// TIA Portal V17 export
FUNCTION "FC_T02_Bobines" : Void   // FC102, LAD
{ S7_Optimized_Access := 'TRUE' }
// stored: SetENOAutomatically false
   VAR_INPUT
      Entree_1 : Bool;
      Bp_Set : Bool;
      Bp_Reset : Bool;
      Entree_2 : Bool;
   END_VAR
   VAR_OUTPUT
      Sortie_1 : Bool;
      Sortie_2 : Bool;
      Sortie_3 : Bool;
   END_VAR
   VAR_IN_OUT
      Memoire : Bool;
   END_VAR
BEGIN

REGION Network 1: Bobine simple
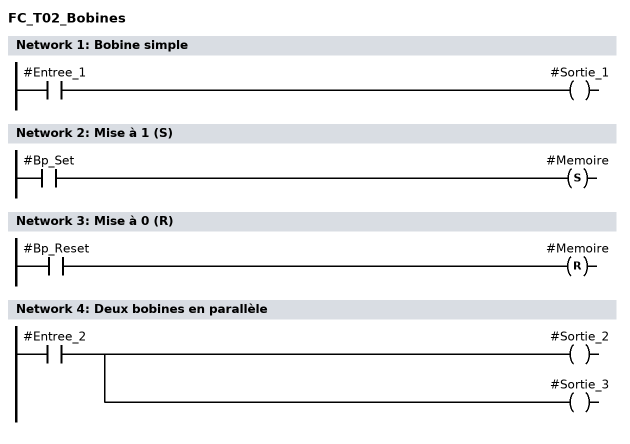
   RUNG wire#powerrail
      Contact( #Entree_1 )
      Coil( #Sortie_1 )
   END_RUNG
   // the same network as SCL:
   #Sortie_1 := #Entree_1;
END_REGION

REGION Network 2: Mise à 1 (S)
   RUNG wire#powerrail
      Contact( #Bp_Set )
      S_Coil( #Memoire )
   END_RUNG
   // the same network as SCL:
   IF #Bp_Set THEN #Memoire := TRUE; END_IF;
END_REGION

REGION Network 3: Mise à 0 (R)
   RUNG wire#powerrail
      Contact( #Bp_Reset )
      R_Coil( #Memoire )
   END_RUNG
   // the same network as SCL:
   IF #Bp_Reset THEN #Memoire := FALSE; END_IF;
END_REGION

REGION Network 4: Deux bobines en parallèle
   RUNG wire#powerrail
      Contact( #Entree_2 )
      wire#w1
      Coil( #Sortie_2 )
   END_RUNG
   RUNG wire#w1
      Coil( #Sortie_3 )
   END_RUNG
   // the same network as SCL:
   #Sortie_2 := #Entree_2;
   #Sortie_3 := #Entree_2;
END_REGION
END_FUNCTION
